(* IEC 61131-3 sources: Palletizer_Control_with_Automation_Studio/Palletizer/Logical/Libraries/AsArLog, 3 files *)

(* ---- AsArLog.typ ---- *)
(********************************************************************
 * COPYRIGHT -- Bernecker + Rainer
 ********************************************************************
 * Library: AsArLog
 * File: AsArLog.typ
 * Author: B+R
 ********************************************************************
 * Data types of library AsArLog
 ********************************************************************)

 TYPE
    asarlogRead : STRUCT
        len             : UDINT;					(*length of the entire log entry (header + binary log data + ASCII string)*)
		lenBin          : UDINT;					(*length of the binary log data*)
		lenAscii        : UDINT;					(*length of the ASCII log data*)
		logLevel        : UDINT;					(*log level of the log entry*)
		errornr         : UDINT;					(*error number of the entry*)
		taskName		: ARRAY[0..35] OF USINT;	(*task name*)
		errYear         : UDINT;					(*year (date of error)*)
		errMonth        : UDINT;					(*month (date of error)*)
		errDay          : UDINT;					(*day (date of error)*)
		errHour         : UDINT;					(*hour (time of error)*)
		errMinute       : UDINT;					(*minute (time of error)*)
		errSecond       : UDINT;					(*second (time of error)*)
		errMilliSec     : UDINT;					(*millisecond (time of error)*)
		errMicroSec     : UDINT;					(*microsecond (time of error)*)
	END_STRUCT;
END_TYPE

(* ---- AsArLog.fun ---- *)
(********************************************************************
 * COPYRIGHT -- Bernecker + Rainer
 ********************************************************************
 * Library: AsArLog
 * File: AsArLog.fun
 * Author: B+R
 ********************************************************************
 * Functions and function blocks of library AsArLog
 ********************************************************************)

 FUNCTION_BLOCK AsArLogCreate					(*creates an AR logger user module; asynchronous execution*)
	VAR_INPUT
		enable		: BOOL;						(*enables execution*)
		pName		: UDINT;					(*name of the AR logger user module to be created give as a pointer, e.g. "vclog".*)
		len     	: UDINT;					(*length of the log data area*)
		memType    	: UDINT;					(*memory type on the target: arlogDRAM, arlogUSRRAM, arlogUSRROM*)
	END_VAR

	VAR
        intResult	: UDINT;					(*internal variable*)
        intState    : UDINT;					(*internal variable*)
        intRes      : UDINT;					(*internal variable*)
	END_VAR

	VAR_OUTPUT
		status		: UINT; 					(*execution status: ERR_OK, ERR_FUB_ENABLE_FALSE, ERR_FUB_BUSY, 0xXXXX = see help*)
		ident		: UDINT;					(*ident of the AR logger basis module to be generated*)
	END_VAR
END_FUNCTION_BLOCK

FUNCTION_BLOCK AsArLogDelete					(*deletes an AR logger user module; asynchronous execution*)
	VAR_INPUT
		enable		: BOOL;						(*enables execution*)
		ident		: UDINT;					(*ident of the AR logger user module to be deleted*)
	END_VAR

	VAR
        intResult	: UDINT;					(*internal variable*)
        intState    : UDINT;					(*internal variable*)
        intRes      : UDINT;					(*internal variable*)
	END_VAR

	VAR_OUTPUT
		status		: UINT; 					(*execution status: ERR_OK, ERR_FUB_ENABLE_FALSE, ERR_FUB_BUSY, 0xXXXX = see help*)
	END_VAR
END_FUNCTION_BLOCK

FUNCTION_BLOCK AsArLogWrite						(*writes a log entry to a AR logger user module; asynchronous execution*)
	VAR_INPUT
		enable		: BOOL;						(*enables execution*)
		ident		: UDINT;					(*ident for the AR logger module to be written (user module or base module)*)
		logLevel	: UDINT;					(*log level of the log entry*)
		errornr		: UDINT;					(*error number of the entry*)
		mem			: UDINT;					(*binary log data given as a pointer*)
		len			: UDINT;					(*length of the binary log data in bytes*)
		asciiString	: UDINT;					(*log-specific zero-terminated ASCII string give as a pointer*)
	END_VAR

	VAR
        intResult	: UDINT;					(*internal variable*)
        intState    : UDINT;					(*internal variable*)
        intRes      : UDINT;					(*internal variable*)
		intTaskName	: ARRAY[0..35] OF USINT;	(*internal variable*)
		intRtkTime  : ARRAY[0..3] OF UDINT;		(*internal variable*)
	END_VAR

	VAR_OUTPUT
		status		: UINT;  					(*execution status: ERR_OK, ERR_FUB_ENABLE_FALSE, ERR_FUB_BUSY, 0xXXXX = see help*)
	END_VAR
END_FUNCTION_BLOCK

FUNCTION_BLOCK AsArLogRead						(*reads a log entry from a AR logger module; asynchronous execution*)
	VAR_INPUT
		enable		: BOOL;						(*enables execution*)
		ident		: UDINT;					(*ident for the AR logger module to be read (user module or base module)*)
		index		: UDINT;					(*index of the log entry to be read*)
		arlogRead	: UDINT;					(*specifies read structure (given as a pointer) where the header data for the log entry can be copied*)
		memBin		: UDINT;					(*buffer for binary log data given as a pointer (if NULL, no binary log data is copied)*)
		lenBin		: UDINT;					(*number of binary log data bytes to be read (if NULL, no binary log data is copied)*)
		memAscii	: UDINT;					(*buffer for ASCII string given as a pointer*)
		lenAscii	: UDINT;					(*number of bytes to be read for the ASCII string*)
	END_VAR

	VAR
        intResult	: UDINT;					(*internal variable*)
        intState    : UDINT;					(*internal variable*)
        intRes      : UDINT;					(*internal variable*)
	END_VAR

	VAR_OUTPUT
		status		: UINT;  					(*execution status: ERR_OK, ERR_FUB_ENABLE_FALSE, ERR_FUB_BUSY, 0xXXXX = see help*)
	END_VAR
END_FUNCTION_BLOCK

FUNCTION_BLOCK AsArLogClear						(*deletes or reinitializes the log data in an AR logger user module; asynchronous execution*)
	VAR_INPUT
		enable		: BOOL;						(*enables execution*)
		ident		: UDINT;					(*ident of the AR logger user module to be reinitialized*)
	END_VAR

	VAR
        intResult	: UDINT;					(*internal variable*)
        intState    : UDINT;					(*internal variable*)
        intRes      : UDINT;					(*internal variable*)
	END_VAR

	VAR_OUTPUT
		status		: UINT; 					(*execution status: ERR_OK, ERR_FUB_ENABLE_FALSE, ERR_FUB_BUSY, 0xXXXX = see help*)
	END_VAR
END_FUNCTION_BLOCK

FUNCTION_BLOCK AsArLogGetInfo					(*reads information from a self-generated AR logger user module or AR logger base user module*)
	VAR_INPUT
		enable		: BOOL;						(*enables execution*)
		pName		: UDINT;					(*name of the AR logger user module (e.g. "vclog") given as a pointer*)
	END_VAR

	VAR
        intResult	: UDINT;					(*internal variable*)
        intState    : UDINT;					(*internal variable*)
        intRes      : UDINT;					(*internal variable*)
	END_VAR

	VAR_OUTPUT
		status		: UINT;						(*execution status: ERR_OK, ERR_FUB_ENABLE_FALSE, 0xXXXX = see help*)
		ident		: UDINT;					(*ident of the AR logger BR module*)
		len	    	: UDINT;					(*length of the log data area*)
		memType		: UDINT;					(*memory type on the target*)
		actualIndex	: UDINT;					(*current entry index in the specified AR logger BR module*)
		FormatVer   : UDINT;					(*version of de log data format*)

	END_VAR
END_FUNCTION_BLOCK

(* ---- AsArLog.var ---- *)
(********************************************************************
 * COPYRIGHT -- Bernecker + Rainer
 ********************************************************************
 * Library: AsArLog
 * File: AsArLog.var
 * Author: B+R
 ********************************************************************
 * Local variables of library AsArLog
 ********************************************************************)

 VAR CONSTANT
	arlogDRAM						 : USINT := 65;		(*temporary AR log modules (DRAM)*)
	arlogUSRRAM						 : USINT := 3;		(*USERRAM*)
	arlogUSRROM						 : USINT := 2;		(*USERROM (USER FLASH)*)

	arlogLEVEL_INFO                  : UDINT := 1;		(*log level INFO*)
	arlogLEVEL_WARNING               : UDINT := 2;		(*log level WARNING*)
	arlogLEVEL_FATAL	             : UDINT := 3;		(*log level FATAL*)

	arlogMIN_LOGDATA_SIZE            : UINT := 4096;	(*minimum log data size of 4 KB*)

	arlogBASE_SYSTEM_LOG_IDENT       : UDINT := 0;		(*fixed ID for the "$arlogsys" base system module*)
	arlogBASE_USER_LOG_IDENT         : UDINT := 1;		(*fixed ID for the "$arlogusr" base user module*)
	arlogBASE_FIELDBUS_LOG_IDENT	 : UDINT := 2;		(*fixed ID for the "fieldbus" logger module*)
	arlogBASE_SAFETY_LOG_IDENT		 : UDINT := 3;		(*fixed ID for the "safety" logger module*)

	arlogERR_ILL_NAME                : UINT := 31400;	(*incorrect or invalid name*)
	arlogERR_ILL_MEMTYPE             : UINT := 31401;	(*incorrect memory type*)
	arlogERR_ILL_LOGLEVEL            : UINT := 31402;	(*invalid log level (only arlogLEVEL_INFO, arlogLEVEL_WARNING, and arlogLEVEL_FATAL valid)*)
	arlogERR_ILL_PARAM               : UINT := 31403;	(*invalid parameters specified*)
	arlogERR_ILL_LEN                 : UINT := 31404;	(*incorrect log data length. Must be >= arlogMIN_LOGDATA_SIZE (4096 bytes)*)
	arlogERR_EXISTING                : UINT := 31405;	(*log module already exists*)
	arlogERR_CREATE                  : UINT := 31406;	(*general create error (create failed)*)
	arlogERR_INSTALL                 : UINT := 31407;	(*install error for AsArLogCreate*)
	arlogERR_ACCESS_DENIED           : UINT := 31408;	(*cannot access the "$arlogsys" and "$arlogusr" base log modules*)
	arlogERR_IN_ACCESS               : UINT := 31409;	(*access denied since other critical FBK simultaneously active*)
	arlogERR_INVALID_IDENT           : UINT := 31410;	(*invalid ident specified*)
	arlogERR_DELETE                  : UINT := 31411;	(*general delete error (delete failed)*)

	arlogERR_NOMEMORY                : UINT := 31412;	(*not enough buffer to copy*)
	arlogERR_NOTEXISTING             : UINT := 31416;	(*AR log module doesn't exist*)

	arlogERR_WRITE                   : UINT := 31417;	(*general write error (write failed)*)
	arlogERR_WRITE_CALC_DATA         : UINT := 31418;	(*error calculating referencing index*)

	arlogERR_READ                    : UINT := 31419;	(*general read error (read failed)*)
	arlogERR_READ_BUFFER             : UINT := 31420;	(*invalid buffer specified*)
	arlogERR_INVALID_INDEX           : UINT := 31421;	(*invalid index (smaller than the reference index and larger than the current index)*)
	arlogERR_INVALID_ENTRY           : UINT := 31422;	(*invalid log entry read*)
	arlogERR_READ_BINARY_BUFFER      : UINT := 31423;	(*buffer length for binary data too small*)
	arlogERR_READ_ASCII_BUFFER       : UINT := 31424;	(*buffer length for ASCII data too small*)
	arlogERR_NO_MORE_ENTRY           : UINT := 31425;	(*FBK still working*)
END_VAR
